(* CODESYS project listof.library
   DefaultNamespace: KOSTAL.AF2024.Core.ListOf
   DocFormat: reStructuredText
   Description: Lists of different elements
   Author: Frank Dümpelmann
   Title: KOSTAL.AF2024.Core.ListOf
   Version: 1.0.0.0
   Company: KOSTAL GmbH & Co.KG
   Placeholder: KOSTAL.AF2024.Core.ListOf

Project tree, tasks and I/O mapping:
  libraries: KOSTAL.AF2024.Core.functionResponse, 0.0.0.2 (KOSTAL GmbH & Co.KG); KOSTAL.AF2024.Core.Settings, 0.0.0.1 (KOSTAL GmbH & Co.KG); KOSTAL.AF2024.Core.System, 0.0.0.1 (KOSTAL GmbH & Co.KG); Tc2_Standard, 3.3.3.0 (Beckhoff Automation GmbH)
  _Interface/
    0_Core/
      BaseElement/
        data type _P_Interface
        data type _ST_Interface
      function block _FB_Interface_Core [ST]: FB_exit, FB_init, _addItem, _findItem, _findItemByIndex, _insertItem, _removeFromBegin, _removeFromEnd, _removeItem, _removeItemByIndex, _nextItem, _previousItem, _clearResult, _setResultFail, _setResultPass, _checkConsistency, _clear, _NumberOfMember, _RegKey
      interface _I_Interface_Core
      interface _I_Interface_Core_Owner
    1_Base/
      function block _FB_Interface_Base [ST]: _verifyMember, _addMember, _findMember, _findMemberByIndex, _insertMember, _removeFromBegin, _removeFromEnd, _removeMember, _removeMemberByIndex, _clear, FB_exit, FB_init
      interface _I_Interface_Base
      interface _I_Interface_Base_Owner
  _Object/
    function block _FB_Object_Base [ST]: _removePayload, _removeMember, _clear, FB_exit, FB_init
    interface _I_Object_Base
    interface _I_Object_Base_Owner
  _STRING/
    0_Core/
      BaseElement/
        data type _P_String
        data type _ST_String
      function block _FB_String_Core [ST]: _addItem, _findItem, _findItemByIndex, _insertItem, _removeFromBegin, _removeFromEnd, _removeItem, _removeItemByIndex, _nextItem, _previousItem, _clearResult, _setResultFail, _setResultPass, _checkConsistency, _clear, _NumberOfMember, FB_exit, FB_init
      interface _I_String_Core
      interface _I_String_Core_Owner
    1_Base/
      function block _FB_String_Base [ST]: _FIFO_peek, _FIFO_pop, _FIFO_push, _addMember, _findMember, _findMemberByIndex, _insertMember, _removeFromBegin, _removeFromEnd, _removeMember, _removeMemberByIndex, _clear, FB_exit, FB_init
      interface _I_String_Base
      interface _I_String_Base_Owner
    function block FB_ListOfString [ST]: addLine, clear, line_GET, line_SET, maxLine, NumberOfLines, removeLine
    interface I_ListOfString: line_GET, maxLine, NumberOfLines
    interface I_ListOfString_Owner: addLine, clear, line_GET, line_SET, maxLine, NumberOfLines, removeLine
  _STRING_UTF8/
    0_Core/
      BaseElement/
        data type P_String_UTF8
        data type ST_String_UTF8
      function block _FB_String_UTF8_Core [ST]: _addItem, _findItem, _findItemByIndex, _insertItem, _removeFromBegin, _removeFromEnd, _removeItem, _removeItemByIndex, _nextItem, _previousItem, _clearResult, _setResultFail, _setResultPass, _checkConsistency, _clear, _NumberOfMember, FB_exit, FB_init
      interface _I_String_UTF8_Core
      interface _I_String_UTF8_Core_Owner
    1_Base/
      function block _FB_String_UTF8_Base [ST]: _FIFO_peek, _FIFO_pop, _FIFO_push, _addMember, _findMember, _findMemberByIndex, _insertMember, _removeFromBegin, _removeFromEnd, _removeMember, _removeMemberByIndex, _clear, FB_exit, FB_init
      interface _I_String_UTF8_Base
      interface _I_String_UTF8_Base_Owner
    function block FB_ListOfString_UTF8 [ST]: addLine, clear, line_GET, line_SET, maxLine, NumberOfLines, removeLine
    interface I_ListOfString_UTF8: line_GET, maxLine, NumberOfLines
    interface I_ListOfString_UTF8_Owner: addLine, clear, line_GET, line_SET, maxLine, NumberOfLines, removeLine
  Project Information/
    function F_GetCompany [ST]
    function F_GetTitle [ST]
    function F_GetVersion [ST]
  Version/
    global variables Global_Version
*)

// _Interface/0_Core/BaseElement/_P_Interface
//Pointer to an element of List
TYPE _P_Interface : POINTER TO _ST_Interface; END_TYPE

// _Interface/0_Core/BaseElement/_ST_Interface
{attribute 'enable_dynamic_creation'}
TYPE _ST_Interface :
	STRUCT
			pNext	 		: _P_Interface;				//Pointer to next Item
			iMember		: KOSTAL_AF2024_Core_System.I_Interface;	//Interface of this item
			pPrevious : _P_Interface;				//Pointer to previous item
	END_STRUCT
END_TYPE

// _STRING/0_Core/BaseElement/_P_String
//Pointer to an element of List
TYPE _P_String : POINTER TO _ST_String; END_TYPE

// _STRING/0_Core/BaseElement/_ST_String
{attribute 'enable_dynamic_creation'}
TYPE _ST_String :
	STRUCT
			pNext	 		: _P_String;														//Pointer to next Item
			Member		: KOSTAL_AF2024_Core_Settings.T_MaxString;	//Text content
			pPrevious : _P_String;														//Pointer to previous item
	END_STRUCT
END_TYPE

// _STRING_UTF8/0_Core/BaseElement/P_String_UTF8
//Pointer to an element of List
TYPE P_String_UTF8 : POINTER TO ST_String_UTF8; END_TYPE

// _STRING_UTF8/0_Core/BaseElement/ST_String_UTF8
{attribute 'enable_dynamic_creation'}
TYPE ST_String_UTF8 :
	STRUCT
			pNext	 		: P_String_UTF8;				//Pointer to next Item
			Member			: KOSTAL_AF2024_Core_Settings.T_MaxString_UTF8;	//Text content
			pPrevious : P_String_UTF8;				//Pointer to previous item
	END_STRUCT
END_TYPE

// Version/Global_Version
{attribute 'TcGenerated'}
{attribute 'no-analysis'}
{attribute 'linkalways'}
// This function has been automatically generated from the project information.
VAR_GLOBAL CONSTANT
	{attribute 'const_non_replaced'}
	stLibVersion_KOSTAL_AF2024_Core_ListOf : ST_LibVersion := (iMajor := 1, iMinor := 0, iBuild := 0, iRevision := 0, nFlags := 0, sVersion := '1.0.0.0');
END_VAR

// _Interface/0_Core/_FB_Interface_Core
(*

| =========================================================================
| List of Items from base Interface {KOSTAL_TC3_Core_System.I_Interface} 
| =========================================================================

..code::

	//In addition to the interface, each item contains the pointer to the previous item 
	//as well as the pointer to the next item in the list.

	TYPE ST_List :
		STRUCT
				pNext			: P_List;
				iMember		: KOSTAL_TC3_Core_System.I_Interface;	
				pPrevious : P_List;
		END_STRUCT
	END_TYPE

============= ======================================= ======================
| The List is defined by (p)Begin and (p)End and also the count of Members 
----------------------------------------------------------------------------
============= ======================================= ======================
 **_pBegin**  >>>>>>>>>>>>>>>>>>>>>>>>>>>>>>>>>>>>>>  **_pEnd**                     
 **Item-1**	    Item-2   Item-3   Item-4  Item-5      **Item-n**                   
============= ======================================= ======================



| =========================================================================
| The Member is an Interface as payload and an access pointer to the        
| previous member and the next member                                      
| ---------------------------------------------------------------------------
| Previous Item ---<<<Pointer-Previous-[Item]-Pointer-Next>>>---NextItem---
| =========================================================================

*)
FUNCTION_BLOCK ABSTRACT _FB_Interface_Core IMPLEMENTS _I_Interface_Core, _I_Interface_Core_Owner

VAR
	_pBegin	: _P_Interface;	//origin of List
  _pEnd		: _P_Interface;	//end of List
	_Count	: UDINT;	//number of registered Member
	
	_RegKeyValue	: UDINT:= UDINT#0;	//use to create an unique ID
	
END_VAR

METHOD FB_exit : BOOL
VAR_INPUT
	bInCopyCode : BOOL; // if TRUE, the exit method is called for exiting an instance that is copied afterwards (online change).
END_VAR

_clear();
END_METHOD

METHOD FB_init : BOOL
VAR_INPUT
	bInitRetains : BOOL; // if TRUE, the retain variables are initialized (warm start / cold start)
	bInCopyCode : BOOL;  // if TRUE, the instance afterwards gets moved into the copy code (online change)
END_VAR

_clear();
END_METHOD

(*
	add new item to end of list
*)
METHOD PROTECTED _addItem : BOOL

VAR_INPUT
	Item		: KOSTAL_AF2024_Core_System.I_Interface;
	Result	: KOSTAL_AF2024_Core_functionResponse.I_T_functionResponse_Owner;
END_VAR

VAR
	_pNewItem	: _P_Interface;
END_VAR

_clearResult(Result);

IF Item = 0 THEN _setResultFail(Result, "Parameter Item is empty");	RETURN;	END_IF


//create a new Item
_pNewItem:= __NEW(_ST_Interface);

//If creation failed 
IF _pNewItem = 0 THEN _setResultFail(Result, "New Item cannot create");	RETURN;	END_IF

//If list is empty
IF THIS^._Count = 0 (*THIS^._pEnd = 0*) THEN THIS^._pBegin:= THIS^._pEnd:= _pNewItem; 
ELSE

	//set new item previous item to actual last item (THIS^._pEnd)
	_pNewItem^.pPrevious:= THIS^._pEnd;
	_pNewItem^.pPrevious^.pNext:= _pNewItem;
 
	THIS^._pEnd:= _pNewItem;
END_IF

THIS^._pEnd^.iMember:= Item;
THIS^._Count:= THIS^._Count + UDINT#1;

_setResultPass(Result, "addItem successful");

_RegKeyValue:= _RegKeyValue + 1;

_addItem:= TRUE;
END_METHOD

(*
	Search for the element {Item} in the list and return {FoundItem} if it is found {_findItem = TRUE}
*)
METHOD PROTECTED _findItem : BOOL
VAR_INPUT
	Item			: KOSTAL_AF2024_Core_System.I_Interface;
	FoundItem	: REFERENCE TO _P_Interface;
	Result		: KOSTAL_AF2024_Core_functionResponse.I_T_functionResponse_Owner;
END_VAR

VAR
	_Item		: _P_Interface;
END_VAR

_clearResult(Result);

IF Item = 0 										THEN _setResultFail(Result, "Parameter Item is empty");	RETURN;	END_IF
IF NOT __ISVALIDREF(FoundItem)	THEN _setResultFail(Result, "FoundItem has no valid reference");	RETURN;	END_IF


_Item := THIS^._pBegin;

WHILE _Item <> 0 DO

	IF _Item^.iMember = Item THEN

		FoundItem := _Item;

		_findItem:= TRUE;

		_setResultPass(Result, "Item found");
		
		RETURN;   

	END_IF
	
	_Item := THIS^._nextItem(_Item, 0);

END_WHILE

//FoundItem:= _Item;

_setResultFail(Result, "Item not found");

_findItem:= FALSE;
END_METHOD

(*
	Search for the element {Item} in the list and return {FoundItem} if it is found {_findItem = TRUE}
*)
METHOD PROTECTED _findItemByIndex : BOOL
VAR_INPUT
	Index			: UDINT;
	FoundItem	: REFERENCE TO _P_Interface;
	Result		: KOSTAL_AF2024_Core_functionResponse.I_T_functionResponse_Owner;
END_VAR

VAR
	_Item		: _P_Interface;
	_udi: UDINT;
END_VAR

_findItemByIndex:= FALSE;

_clearResult(Result);

IF _Count = 0										THEN _setResultFail(Result, "List is empty");											RETURN;	END_IF
IF Index > (_Count - 1)					THEN _setResultFail(Result, "Parameter Index is out of range");		RETURN;	END_IF
IF NOT __ISVALIDREF(FoundItem)	THEN _setResultFail(Result, "FoundItem has no valid reference");	RETURN;	END_IF

//set index 0
_Item := THIS^._pBegin;

//increase until index is reached
FOR _udi:= 1 TO Index DO
		_Item := THIS^._nextItem(_Item, 0);
END_FOR

FoundItem:= _Item;

IF FoundItem = 0 THEN
	_setResultFail(Result, "Item not found");
ELSE	
	_setResultPass(Result, "Item found");
	_findItemByIndex:= TRUE;
END_IF
END_METHOD

METHOD PROTECTED _insertItem : BOOL
VAR_INPUT
	Index		: UDINT;	//Index a which shall inserted the {Item}
	Item		: KOSTAL_AF2024_Core_System.I_Interface;
	Result		: KOSTAL_AF2024_Core_functionResponse.I_T_functionResponse_Owner;
END_VAR

VAR
	_pNewItem			: _P_Interface;
	_pExitingItem	: _P_Interface;
END_VAR

_clearResult(Result);

//Item is empty
IF Item = 0 THEN _setResultFail(Result, "Parameter Item is empty");	RETURN;	END_IF

//if List is empty add item 
IF (Index = 0) AND (_Count = 0)	THEN _insertItem:= _addItem(Item, Result);	RETURN;	END_IF

//Index is in list not available 
IF Index > (_Count - 1) THEN _setResultFail(Result, "Index is out of range");	RETURN;	END_IF

//if index is end of list then add item to end of list 
IF (Index = (_Count - 1)) THEN _insertItem:= _addItem(Item, Result);	RETURN;	END_IF

//try to find item where shall inserted
IF NOT _findItemByIndex(Index, _pExitingItem, Result) THEN RETURN;	END_IF
IF _pExitingItem = 0 THEN _setResultFail(Result, "Item not available");	RETURN;	END_IF


//create a new Item
_pNewItem:= __NEW(_ST_Interface);

//If creation failed 
IF _pNewItem = 0 THEN _setResultFail(Result, "New Item cannot create");	RETURN;	END_IF

_pNewItem^.iMember:= Item;

_pNewItem^.pNext		:= _pExitingItem;							//set the next item from new item to existing founded item
_pNewItem^.pPrevious:= _pExitingItem^.pPrevious;	//set the previous from existing item to the previous of new item

//if a previous exist then
//set the next from previous from existing item to the previous of new item
IF _pNewItem^.pPrevious <> 0 THEN	_pNewItem^.pPrevious^.pNext:= _pNewItem;	END_IF

_pExitingItem^.pPrevious:= _pNewItem;							//set the previous from existing founded item to  new item

//if inserted at the begin of list, set the begin pointer to new Item
IF _pBegin = _pExitingItem THEN	_pBegin:= _pNewItem;	END_IF

_Count:= _Count + UDINT#1;

_setResultPass(Result, "insertItem successful");

_RegKeyValue:= _RegKeyValue + 1;

_insertItem:= TRUE;
END_METHOD

(*
	remove Item from begin of list
*)
METHOD PROTECTED _removeFromBegin : BOOL
VAR_INPUT
	Result	: KOSTAL_AF2024_Core_functionResponse.I_T_functionResponse_Owner;
END_VAR

_removeFromBegin:= _removeItemByIndex(0, Result);
END_METHOD

(*
	remove Item from end of list
*)
METHOD PROTECTED _removeFromEnd : BOOL
VAR_INPUT
	Result	: KOSTAL_AF2024_Core_functionResponse.I_T_functionResponse_Owner;
END_VAR

_removeFromEnd:= _removeItemByIndex(_Count - 1, Result);
END_METHOD

(*
	remove given {Item} from List
*)
METHOD PROTECTED _removeItem : BOOL
VAR_INPUT
	Item		: _P_Interface;
	Result	: KOSTAL_AF2024_Core_functionResponse.I_T_functionResponse_Owner;
END_VAR

_clearResult(Result);

IF Item = 0 THEN _setResultFail(Result, "Parameter Item is empty");	RETURN;	END_IF

//exist a next member
IF Item^.pNext <> 0 THEN
	//set next members previous Item  to my previous Item
	Item^.pNext^.pPrevious := Item^.pPrevious; 
END_IF

//exist a previous member
IF Item^.pPrevious <> 0 THEN
	//set previous members next Item  to my next Item
	Item^.pPrevious^.pNext := Item^.pNext;
END_IF

//Item is the once member
IF Item = _pBegin AND Item = _pEnd THEN
	
	_pBegin := 0;
	_pEnd := 0;

ELSIF Item = _pBegin (*AND Item <> THIS^._pEnd*) THEN

	_pBegin := Item^.pNext;

ELSIF Item = _pEnd THEN

	_pEnd := Item^.pPrevious;

END_IF

__DELETE(Item);

IF  _Count > UDINT#0 THEN	_Count := _Count - UDINT#1;	
ELSE
	_setResultFail(Result, "removeItem Counter underflow");
	RETURN;
END_IF

_setResultPass(Result, "removeItem successful");
_removeItem:= TRUE;
END_METHOD

(*
	remove given {Index} from List
*)
METHOD PROTECTED _removeItemByIndex : BOOL
VAR_INPUT
	Index		: UDINT;
	Result	: KOSTAL_AF2024_Core_functionResponse.I_T_functionResponse_Owner;
END_VAR

VAR
	_Item		: _P_Interface;
	_bFound	: BOOL;
END_VAR

IF NOT _findItemByIndex(Index, _Item, Result)	THEN RETURN;	END_IF

_removeItemByIndex:= _removeItem(_Item, Result);
END_METHOD

// retreives the pointer to the next item of the given entry
METHOD PROTECTED _nextItem : _P_Interface;
VAR_INPUT
    Item : _P_Interface;
		Result	: KOSTAL_AF2024_Core_functionResponse.I_T_functionResponse_Owner;
END_VAR
VAR
	_Res	: _P_Interface;
END_VAR

IF Item <> 0 THEN	_Res := Item^.pNext;
ELSE							_Res := 0;
END_IF

_nextItem:= _Res;
END_METHOD

// retreives the previous item of the given entry
METHOD PROTECTED _previousItem : _P_Interface
VAR_INPUT
    Item 	: _P_Interface;
END_VAR
VAR
	_Res	: _P_Interface;
END_VAR

IF Item <> 0 THEN	_Res := Item^.pPrevious;
ELSE							_Res := 0;
END_IF

_previousItem:= _Res;
END_METHOD

(*
	Clear result component
*)
METHOD PROTECTED _clearResult : BOOL
VAR_INPUT
	IN : KOSTAL_AF2024_Core_functionResponse.I_T_functionResponse_Owner;
END_VAR

IF IN <> 0 THEN  
	 IN.clear();
	_clearResult:= TRUE;	
END_IF
END_METHOD

(*
	set result to fail with given information 
*)
METHOD PROTECTED _setResultFail : BOOL
VAR_INPUT
	IN 		: KOSTAL_AF2024_Core_functionResponse.I_T_functionResponse_Owner;
	Info	: KOSTAL_AF2024_Core_Settings.T_MaxString;
END_VAR

IF IN <> 0 THEN 

	IN.success:= FALSE;
	IN.status:= Info;

	_setResultFail:= TRUE;

END_IF
END_METHOD

(*
	set result to pass with given information 
*)
METHOD PROTECTED _setResultPass : BOOL
VAR_INPUT
	IN 		: KOSTAL_AF2024_Core_functionResponse.I_T_functionResponse_Owner;
	Info	: KOSTAL_AF2024_Core_Settings.T_MaxString;
END_VAR

IF IN <> 0 THEN 

	IN.success:= TRUE;
	IN.status:= Info;

	_setResultPass:= TRUE;

END_IF
END_METHOD

(*
	Check if the list is consistent
*)
METHOD PROTECTED _checkConsistency : BOOL
VAR_INPUT
	Result	: KOSTAL_AF2024_Core_functionResponse.I_T_functionResponse_Owner;
END_VAR

VAR
	_pItem			: _P_Interface;
	_pNext			: _P_Interface;
	_pPrev			: _P_Interface;
	_nItemCounter	: UDINT;
	_bBeginOk			: BOOL;
	_bEndOk			: BOOL;
	_bPrevLinkOk		: BOOL;
	_bNextLinkOk		: BOOL;
	_bItemCountOk	: BOOL;
	_bInterfaceOk	: BOOL;
END_VAR

// check from pHead to pTail
_pItem:= _pBegin;
_nItemCounter:= 0;

IF _pBegin <> 0 THEN
	_bBeginOk:= (_pBegin^.pPrevious = 0);
ELSE
	_bBeginOk:= TRUE;
END_IF

IF _pEnd <> 0 THEN
	_bEndOk:= (_pEnd^.pNext = 0);
ELSE
	_bEndOk:= TRUE;
END_IF

IF _bBeginOk AND _bEndOk THEN

	_bPrevLinkOk:= TRUE;
	_bNextLinkOk:= TRUE;
	_bInterfaceOk:= TRUE;

	WHILE _pItem <> 0 DO
		
		_pPrev:= _pItem^.pPrevious;
		_pNext:= _pItem^.pNext;

		IF _pPrev <> 0 THEN
			_bPrevLinkOk:= (_pPrev^.pNext = _pItem);
		ELSE
			_bPrevLinkOk:= (_pItem = _pBegin);
		END_IF

		IF _pNext <> 0 THEN
			_bNextLinkOk:= (_pNext^.pPrevious = _pItem);
		ELSE
			_bNextLinkOk:= (_pItem = _pEnd);
		END_IF

		_bInterfaceOk:= (_pItem^.iMember <> 0);

		IF NOT _bNextLinkOk OR NOT _bPrevLinkOk OR NOT _bInterfaceOk THEN	EXIT;	END_IF

		//handle iteration
		_nItemCounter:= _nItemCounter + UDINT#1;
		_pItem:= _nextItem(_pItem, 0);

	END_WHILE

END_IF

_bItemCountOk:= (_nItemCounter = THIS^._Count);

IF 		NOT _bBeginOk			THEN	_setResultFail(Result, "List head not ok");
ELSIF NOT _bEndOk				THEN	_setResultFail(Result, "List End not ok");
ELSIF NOT _bPrevLinkOk 	THEN	_setResultFail(Result, Tc2_Standard.WCONCAT("Previous Link failed by item ", UDINT_TO_WSTRING(_nItemCounter)));
ELSIF NOT _bNextLinkOk	THEN	_setResultFail(Result, Tc2_Standard.WCONCAT("Next Link failed by item ", UDINT_TO_WSTRING(_nItemCounter)));
ELSIF NOT	_bInterfaceOk	THEN	_setResultFail(Result, Tc2_Standard.WCONCAT("Interface failed by item ", UDINT_TO_WSTRING(_nItemCounter))); 
ELSIF NOT	_bItemCountOk THEN	_setResultFail(Result, "Itemcounter is not ok");
ELSE													_setResultPass(Result, "List is consistent");	_checkConsistency:= TRUE;
END_IF
END_METHOD

(*
	Delete the complete content of the list
*)
METHOD PROTECTED _clear

WHILE THIS^._pBegin <> 0 DO
    THIS^._removeItem(THIS^._pBegin, 0);  
END_WHILE
END_METHOD

//return the nnumber of items in List
PROPERTY PROTECTED _NumberOfMember : UDINT
GET

_NumberOfMember:= _Count;
END_GET
END_PROPERTY

PROPERTY PROTECTED _RegKey : UDINT
GET

_RegKey:= THIS^._RegKeyValue;
END_GET
END_PROPERTY

END_FUNCTION_BLOCK

// _Interface/0_Core/_I_Interface_Core
INTERFACE _I_Interface_Core EXTENDS KOSTAL_AF2024_Core_System.I_Interface

END_INTERFACE

// _Interface/0_Core/_I_Interface_Core_Owner
INTERFACE _I_Interface_Core_Owner EXTENDS KOSTAL_AF2024_Core_System.I_Interface

END_INTERFACE

// _Interface/1_Base/_FB_Interface_Base
(*

| =========================================================================
| List of Items from base Interface {KOSTAL_TC3_Core_System.I_Interface} 
| =========================================================================

..code::

	//In addition to the interface, each item contains the pointer to the previous item 
	//as well as the pointer to the next item in the list.

	TYPE ST_List :
		STRUCT
				pNext			: P_List;
				iMember		: KOSTAL_TC3_Core_System.I_Interface;	
				pPrevious : P_List;
		END_STRUCT
	END_TYPE

============= ======================================= ======================
| The List is defined by (p)Begin and (p)End and also the count of Members 
----------------------------------------------------------------------------
============= ======================================= ======================
 **_pBegin**  >>>>>>>>>>>>>>>>>>>>>>>>>>>>>>>>>>>>>>  **_pEnd**                     
 **Item-1**	    Item-2   Item-3   Item-4  Item-5      **Item-n**                   
============= ======================================= ======================



| =========================================================================
| The Member is an Interface as payload and an access pointer to the        
| previous member and the next member                                      
| ---------------------------------------------------------------------------
| Previous Item ---<<<Pointer-Previous-[Item]-Pointer-Next>>>---NextItem---
| =========================================================================

*)
FUNCTION_BLOCK ABSTRACT _FB_Interface_Base EXTENDS _FB_Interface_Core IMPLEMENTS _I_Interface_Base, _I_Interface_Base_Owner

(*
	integrate here the veryfing of your interface type 
	only if verifing is passed [_verifyMember:= TRUE] the called metode will proceeded 
*)
METHOD PROTECTED _verifyMember : BOOL

VAR_INPUT
	Member	: KOSTAL_AF2024_Core_System.I_Interface;
	Result	: KOSTAL_AF2024_Core_functionResponse.I_T_functionResponse_Owner;
END_VAR

VAR
	_obj	: KOSTAL_AF2024_Core_System.I_Interface;
	_bResult: BOOL;
END_VAR

IF Member = 0 THEN _setResultFail(Result, "Parameter Member is empty");	RETURN;	END_IF

_bResult:= __QUERYINTERFACE(Member, _obj);

IF NOT _bResult OR (_obj = 0) THEN
	IF Result <> 0 THEN  
		Result.success:= FALSE; 
		Result.status:= "no valid interface found";	
	END_IF	
	RETURN;
END_IF

_verifyMember:= TRUE;
END_METHOD

(*
	add new Member to end of list
*)
METHOD PROTECTED _addMember : BOOL

VAR_INPUT
	Member		: KOSTAL_AF2024_Core_System.I_Interface;
	Result	: KOSTAL_AF2024_Core_functionResponse.I_T_functionResponse_Owner;
END_VAR


VAR
	_Member: KOSTAL_AF2024_Core_System.I_Interface;
END_VAR

//IF NOT _verifyMember(Member, Result)	THEN	RETURN;	END_IF

//member already exist
IF _findMember(Member,_Member, Result) THEN 
	_setResultFail(Result, "The participant already exists in the list.");
	RETURN;	
END_IF	

_addMember:= _addItem(Member, Result);
END_METHOD

(*
	Search for the element {Item} in the list and return {FoundItem} if it is found {_findItem = TRUE}
*)
METHOD PROTECTED _findMember : BOOL
VAR_INPUT
	Member			: KOSTAL_AF2024_Core_System.I_Interface;
	FoundMember	: REFERENCE TO KOSTAL_AF2024_Core_System.I_Interface;	//return value
	Result			: KOSTAL_AF2024_Core_functionResponse.I_T_functionResponse_Owner;
END_VAR

VAR
	_Item		: _P_Interface;
END_VAR

_clearResult(Result);

IF Member = 0 												THEN _setResultFail(Result, "Parameter Item is empty");	RETURN;	END_IF
IF NOT __ISVALIDREF(FoundMember)			THEN _setResultFail(Result, "FoundItem has no valid reference");	RETURN;	END_IF
IF NOT _verifyMember(Member, Result)	THEN	RETURN;	END_IF

_findMember:= _findItem(Member, _Item, Result);

IF NOT _findMember		THEN	RETURN;	END_IF
IF _Item = 0 					THEN	RETURN;	END_IF
//IF _Item^.iMember = 0 THEN	RETURN;	END_IF
IF NOT _verifyMember(_Item^.iMember, Result)	THEN	RETURN;	END_IF

FoundMember:= _Item^.iMember;
END_METHOD

//find a modul by index  
METHOD PROTECTED _findMemberByIndex : BOOL
VAR_INPUT
	Index				: UDINT;	//index of item
	FoundMember	: REFERENCE TO KOSTAL_AF2024_Core_System.I_Interface;	//return value
	Result			: KOSTAL_AF2024_Core_functionResponse.I_T_functionResponse_Owner;	//result information
END_VAR

VAR
	_FoundItem	: _P_Interface;
END_VAR

IF NOT __ISVALIDREF(FoundMember)	THEN _setResultFail(Result, "FoundMember has no valid reference");	RETURN;	END_IF

FoundMember:= 0;

_findMemberByIndex:= _findItemByIndex(Index,_FoundItem, Result);

IF NOT _findMemberByIndex THEN RETURN;	END_IF

IF NOT _verifyMember(_FoundItem^.iMember, Result) THEN RETURN;	END_IF

FoundMember:= _FoundItem^.iMember;

_findMemberByIndex:= TRUE;
END_METHOD

METHOD PROTECTED _insertMember : BOOL
VAR_INPUT
	Index		: UDINT;	//Index a which shall inserted the {Item}
	Member	: KOSTAL_AF2024_Core_System.I_Interface;
	Result	:KOSTAL_AF2024_Core_functionResponse.I_T_functionResponse_Owner;
END_VAR

VAR
	_Member: KOSTAL_AF2024_Core_System.I_Interface;
END_VAR

//IF NOT _verifyMember(Member, Result)	THEN	RETURN;	END_IF

//member already exist
IF _findMember(Member,_Member, Result) THEN 
	_setResultFail(Result, "The participant already exists in the list.");
	RETURN;	
END_IF	

_insertMember:= _insertItem(Index, Member, Result);
END_METHOD

(*
	remove Item from begin of list
*)
METHOD PROTECTED _removeFromBegin : BOOL
VAR_INPUT
	Result	: KOSTAL_AF2024_Core_functionResponse.I_T_functionResponse_Owner;
END_VAR

_removeFromBegin:= _removeMemberByIndex(0, Result);
END_METHOD

(*
	remove Item from end of list
*)
METHOD PROTECTED _removeFromEnd : BOOL
VAR_INPUT
	Result	: KOSTAL_AF2024_Core_functionResponse.I_T_functionResponse_Owner;
END_VAR

_removeFromEnd:= _removeMemberByIndex(_Count - 1, Result);
END_METHOD

(*
	remove given {Member} from List
*)
METHOD PROTECTED _removeMember : BOOL
VAR_INPUT
	Member	: KOSTAL_AF2024_Core_System.I_Interface;
	Result	: KOSTAL_AF2024_Core_functionResponse.I_T_functionResponse_Owner;
END_VAR

VAR
	_Item		: _P_Interface;
	_bFound: BOOL;
END_VAR


IF NOT _verifyMember(Member, Result)	THEN	RETURN;	END_IF

_bFound:= _findItem(Member, _Item, Result);

IF NOT _bFound THEN RETURN;	END_IF

_removeMember:= _removeItem(_Item, Result);
END_METHOD

(*
	remove given {Index} from List
*)
METHOD PROTECTED _removeMemberByIndex : BOOL
VAR_INPUT
	Index		: UDINT;
	Result	: KOSTAL_AF2024_Core_functionResponse.I_T_functionResponse_Owner;
END_VAR

VAR
	_bFound	: BOOL;
	_Member	: KOSTAL_AF2024_Core_System.I_Interface;

END_VAR

IF NOT _findMemberByIndex(Index, _Member, Result)	THEN RETURN;	END_IF

_removeMemberByIndex:= _removeMember(_Member, Result);
END_METHOD

(*
	Delete the complete content of the list
*)
METHOD PROTECTED _clear
VAR_INPUT
END_VAR

WHILE THIS^._pBegin <> 0 DO
    THIS^._removeMember(THIS^._pBegin^.iMember, 0);  
END_WHILE
END_METHOD

METHOD FB_exit : BOOL
VAR_INPUT
	bInCopyCode : BOOL; // if TRUE, the exit method is called for exiting an instance that is copied afterwards (online change).
END_VAR

_clear();
END_METHOD

METHOD FB_init : BOOL
VAR_INPUT
	bInitRetains : BOOL; // if TRUE, the retain variables are initialized (warm start / cold start)
	bInCopyCode : BOOL;  // if TRUE, the instance afterwards gets moved into the copy code (online change)
END_VAR

_clear();
END_METHOD

END_FUNCTION_BLOCK

// _Interface/1_Base/_I_Interface_Base
INTERFACE _I_Interface_Base EXTENDS _I_Interface_Core

END_INTERFACE

// _Interface/1_Base/_I_Interface_Base_Owner
INTERFACE _I_Interface_Base_Owner EXTENDS _I_Interface_Core_Owner

END_INTERFACE

// _Object/_FB_Object_Base
(*

| ==================================================================================
| List of Items of objects with base Interface {KOSTAL_TC3_Core_System.I_Interface} 
| ==================================================================================

..code::

	//In addition to the interface, each item contains the pointer to the previous item 
	//as well as the pointer to the next item in the list.

	TYPE ST_List :
		STRUCT
				pNext			: P_List;
				iMember		: KOSTAL_TC3_Core_System.I_Interface;	
				pPrevious : P_List;
		END_STRUCT
	END_TYPE

============= ======================================= ======================
| The List is defined by (p)Begin and (p)End and also the count of Members 
----------------------------------------------------------------------------
============= ======================================= ======================
 **_pBegin**  >>>>>>>>>>>>>>>>>>>>>>>>>>>>>>>>>>>>>>  **_pEnd**                     
 **Item-1**	    Item-2   Item-3   Item-4  Item-5      **Item-n**                   
============= ======================================= ======================



| =========================================================================
| The Member is an object which implements the base Interface as payload. 
| -------------------------------------------------------------------------
| Previous Item ---<<<Pointer-Previous-[Item]-Pointer-Next>>>---NextItem---
| =========================================================================

*)
FUNCTION_BLOCK ABSTRACT _FB_Object_Base EXTENDS _FB_Interface_Base IMPLEMENTS _I_Object_Base, _I_Object_Base_Owner

(*
	Integrate the type-specific procedures here to clean up the member and remove it from memory. 
	only if verifing is passed [_verifyMember:= TRUE] the called metode should proceed 
*)
METHOD PROTECTED _removePayload : BOOL
VAR_INPUT
	Member	: KOSTAL_AF2024_Core_System.I_Interface;
	Result	: KOSTAL_AF2024_Core_functionResponse.I_T_functionResponse_Owner;
END_VAR

_removePayload:= TRUE;
END_METHOD

(*
	remove given {Member} from List including the customer payload {_removePayload()]
*)
METHOD PROTECTED _removeMember : BOOL
VAR_INPUT
	Member	: KOSTAL_AF2024_Core_System.I_Interface;
	Result	: KOSTAL_AF2024_Core_functionResponse.I_T_functionResponse_Owner;
END_VAR

VAR
	_Item		: _P_Interface;
	_bFound: BOOL;
END_VAR

IF NOT _verifyMember(Member, Result)	THEN	RETURN;	END_IF

_bFound:= _findItem(Member, _Item, Result);

IF NOT _bFound THEN RETURN;	END_IF

_removePayload(Member, Result);

_removeMember:= _removeItem(_Item, Result);
END_METHOD

(*
	Delete the complete content of the list including the customer payload {_removePayload()}
*)
METHOD PROTECTED _clear

WHILE THIS^._pBegin <> 0 DO
  _removeMember(_pBegin^.iMember, 0);  
END_WHILE
END_METHOD

METHOD FB_exit : BOOL
VAR_INPUT
	bInCopyCode : BOOL; // if TRUE, the exit method is called for exiting an instance that is copied afterwards (online change).
END_VAR

_clear();
END_METHOD

METHOD FB_init : BOOL
VAR_INPUT
	bInitRetains : BOOL; // if TRUE, the retain variables are initialized (warm start / cold start)
	bInCopyCode : BOOL;  // if TRUE, the instance afterwards gets moved into the copy code (online change)
END_VAR

_clear();
END_METHOD

END_FUNCTION_BLOCK

// _Object/_I_Object_Base
INTERFACE _I_Object_Base EXTENDS _I_Interface_Base

END_INTERFACE

// _Object/_I_Object_Base_Owner
INTERFACE _I_Object_Base_Owner EXTENDS _I_Interface_Base_Owner

END_INTERFACE

// _STRING/0_Core/_FB_String_Core
(*

| =========================================================================
| List of Items from base Interface {KOSTAL_TC3_Core_System.I_Interface} 
| =========================================================================

..code::

	//In addition to the interface, each item contains the pointer to the previous item 
	//as well as the pointer to the next item in the list.

	TYPE ST_List :
		STRUCT
				pNext			: P_List;
				iMember		: KOSTAL_TC3_Core_System.I_Interface;	
				pPrevious : P_List;
		END_STRUCT
	END_TYPE

============= ======================================= ======================
| The List is defined by (p)Begin and (p)End and also the count of Members 
----------------------------------------------------------------------------
============= ======================================= ======================
 **_pBegin**  >>>>>>>>>>>>>>>>>>>>>>>>>>>>>>>>>>>>>>  **_pEnd**                     
 **Item-1**	    Item-2   Item-3   Item-4  Item-5      **Item-n**                   
============= ======================================= ======================



| =========================================================================
| The Member is an Interface as payload and an access pointer to the        
| previous member and the next member                                      
| ---------------------------------------------------------------------------
| Previous Item ---<<<Pointer-Previous-[Item]-Pointer-Next>>>---NextItem---
| =========================================================================

*)
FUNCTION_BLOCK ABSTRACT _FB_String_Core IMPLEMENTS _I_String_Core, _I_String_Core_Owner

VAR
	_pBegin	: _P_String;	//origin of List
  _pEnd		: _P_String;	//end of List
	_Count	: UDINT;	//number of registered Member
END_VAR

(*
	add new item to end of list
*)
METHOD PROTECTED _addItem : BOOL

VAR_INPUT
	Member	: KOSTAL_AF2024_Core_Settings.T_MaxString;
	Result	: KOSTAL_AF2024_Core_functionResponse.I_T_functionResponse_Owner;
END_VAR

VAR
	_pNewItem	: _P_String;
END_VAR

_clearResult(Result);

//IF Item = 0 THEN _setResultFail(Result, 'Parameter Item is empty');	RETURN;	END_IF


//create a new Item
_pNewItem:= __NEW(_ST_String);

//If creation failed 
IF _pNewItem = 0 THEN _setResultFail(Result, "New Item cannot create");	RETURN;	END_IF

//If list is empty
IF _Count = 0 THEN _pBegin:= _pEnd:= _pNewItem; 
ELSE

	//set new item previous item to actual last item (THIS^._pEnd)
	_pNewItem^.pPrevious:= _pEnd;
	_pNewItem^.pPrevious^.pNext:= _pNewItem;
 
	_pEnd:= _pNewItem;

END_IF

_pEnd^.Member:= Member;
_Count:= _Count + UDINT#1;

_setResultPass(Result, "addItem successful");

_addItem:= TRUE;
END_METHOD

(*
	Search for the element {Item} in the list and return {FoundItem} if it is found {_findItem = TRUE}
*)
METHOD PROTECTED _findItem : BOOL
VAR_INPUT
	Member		: KOSTAL_AF2024_Core_Settings.T_MaxString;
	FoundItem	: REFERENCE TO _P_String;
	Result		: KOSTAL_AF2024_Core_functionResponse.I_T_functionResponse_Owner;
END_VAR

VAR
	_Item		: _P_String;
END_VAR

_clearResult(Result);

IF NOT __ISVALIDREF(FoundItem)	THEN _setResultFail(Result, "FoundItem has no valid reference");	RETURN;	END_IF


_Item := _pBegin;

WHILE _Item <> 0 DO

	IF _Item^.Member = Member THEN

		FoundItem := _Item;

		_findItem:= TRUE;

		_setResultPass(Result, "Item found");
		
		RETURN;   

	END_IF
	
	_Item := _nextItem(_Item, 0);

END_WHILE

//FoundItem:= _Item;

_setResultFail(Result, "Item not found");

_findItem:= FALSE;
END_METHOD

(*
	Search for the element {Item} in the list and return {FoundItem} if it is found {_findItem = TRUE}
*)
METHOD PROTECTED _findItemByIndex : BOOL
VAR_INPUT
	Index			: UDINT;
	FoundItem	: REFERENCE TO _P_String;
	Result		: KOSTAL_AF2024_Core_functionResponse.I_T_functionResponse_Owner;
END_VAR

VAR
	_Item	: _P_String;
	_udi	: UDINT;
END_VAR

_findItemByIndex:= FALSE;

_clearResult(Result);

IF _Count = 0										THEN _setResultFail(Result, "List is empty");											RETURN;	END_IF
IF Index > (_Count - 1)					THEN _setResultFail(Result, "Parameter Index is out of range");		RETURN;	END_IF
IF NOT __ISVALIDREF(FoundItem)	THEN _setResultFail(Result, "FoundItem has no valid reference");	RETURN;	END_IF


_Item := _pBegin;

FOR _udi:= 1 TO Index DO
		_Item := _nextItem(_Item, 0);
END_FOR

FoundItem:= _Item;

IF FoundItem = 0 THEN
	_setResultFail(Result, "Item not found");
ELSE	
	_setResultPass(Result, "Item found");
	_findItemByIndex:= TRUE;
END_IF
END_METHOD

METHOD PROTECTED _insertItem : BOOL
VAR_INPUT
	Index		: UDINT;	//Index a which shall inserted the {Item}
	Member	: KOSTAL_AF2024_Core_Settings.T_MaxString;
	Result	: KOSTAL_AF2024_Core_functionResponse.I_T_functionResponse_Owner;
END_VAR

VAR
	_pNewItem			: _P_String;
	_pExitingItem	: _P_String;
END_VAR
_clearResult(Result);

//if List is empty add item 
IF (Index = 0) AND (_Count = 0)	THEN _insertItem:= _addItem(Member, Result);	RETURN;	END_IF

//Index is in list not available 
IF Index > (_Count - 1) THEN _setResultFail(Result, "Index is out of range");	RETURN;	END_IF

//if index is end of list then add item to end of list 
IF (Index = (_Count - 1)) THEN _insertItem:= _addItem(Member, Result);	RETURN;	END_IF

//try to find item where shall inserted
IF NOT _findItemByIndex(Index, _pExitingItem, Result) THEN RETURN;	END_IF
IF _pExitingItem = 0 THEN _setResultFail(Result, "Item not available");	RETURN;	END_IF


//create a new Item
_pNewItem:= __NEW(_ST_String);

//If creation failed 
IF _pNewItem = 0 THEN _setResultFail(Result, "New Item cannot create");	RETURN;	END_IF

_pNewItem^.Member:= Member;

_pNewItem^.pNext		:= _pExitingItem;							//set the next item from new item to existing founded item
_pNewItem^.pPrevious:= _pExitingItem^.pPrevious;	//set the previous from existing item to the previous of new item

//if a previous exist then
//set the next from previous from existing item to the previous of new item
IF _pNewItem^.pPrevious <> 0 THEN	_pNewItem^.pPrevious^.pNext:= _pNewItem;	END_IF

_pExitingItem^.pPrevious:= _pNewItem;							//set the previous from existing founded item to  new item

//if inserted at the begin of list, set the begin pointer to new Item
IF _pBegin = _pExitingItem THEN	_pBegin:= _pNewItem;	END_IF

_Count:= _Count + UDINT#1;

_setResultPass(Result, "insertItem successful");

_insertItem:= TRUE;
END_METHOD

(*
	remove Item from begin of list
*)
METHOD PROTECTED _removeFromBegin : BOOL
VAR_INPUT
	Result	: KOSTAL_AF2024_Core_functionResponse.I_T_functionResponse_Owner;
END_VAR

_removeFromBegin:= _removeItemByIndex(0, Result);
END_METHOD

(*
	remove Item from end of list
*)
METHOD PROTECTED _removeFromEnd : BOOL
VAR_INPUT
	Result	: KOSTAL_AF2024_Core_functionResponse.I_T_functionResponse_Owner;
END_VAR

_removeFromEnd:= _removeItemByIndex(_Count - 1, Result);
END_METHOD

(*
	remove given {Item} from List
*)
METHOD PROTECTED _removeItem : BOOL
VAR_INPUT
	Item		: _P_String;
	Result	: KOSTAL_AF2024_Core_functionResponse.I_T_functionResponse_Owner;
END_VAR

_clearResult(Result);

IF Item = 0 THEN _setResultFail(Result, "Parameter Item is empty");	RETURN;	END_IF

//exist a next member
IF Item^.pNext <> 0 THEN
	//set next members previous Item  to my previous Item
	Item^.pNext^.pPrevious := Item^.pPrevious; 
END_IF

//exist a previous member
IF Item^.pPrevious <> 0 THEN
	//set previous members next Item  to my next Item
	Item^.pPrevious^.pNext := Item^.pNext;
END_IF

//Item is the once member
IF Item = _pBegin AND Item = _pEnd THEN
	
	_pBegin := 0;
	_pEnd := 0;

ELSIF Item = _pBegin THEN

	_pBegin := Item^.pNext;

ELSIF Item = _pEnd THEN

	_pEnd := Item^.pPrevious;

END_IF

__DELETE(Item);

IF  _Count > UDINT#0 THEN	_Count := _Count - UDINT#1;	
ELSE
	_setResultFail(Result, "removeItem Counter underflow");
	RETURN;
END_IF

_setResultPass(Result, "removeItem successful");
_removeItem:= TRUE;
END_METHOD

(*
	remove given {Index} from List
*)
METHOD PROTECTED _removeItemByIndex : BOOL
VAR_INPUT
	Index		: UDINT;
	Result	: KOSTAL_AF2024_Core_functionResponse.I_T_functionResponse_Owner;
END_VAR

VAR
	_Item		: _P_String;
	_bFound	: BOOL;
END_VAR

IF NOT _findItemByIndex(Index, _Item, Result)	THEN RETURN;	END_IF

_removeItemByIndex:= _removeItem(_Item, Result);
END_METHOD

// retreives the pointer to the next item of the given entry
METHOD PROTECTED _nextItem : _P_String;
VAR_INPUT
    Item : _P_String;
		Result	: KOSTAL_AF2024_Core_functionResponse.I_T_functionResponse_Owner;
END_VAR
VAR
	_Res	: _P_String;
END_VAR

IF Item <> 0 THEN	_Res := Item^.pNext;
ELSE							_Res := 0;
END_IF

_nextItem:= _Res;
END_METHOD

// retreives the previous item of the given entry
METHOD PROTECTED _previousItem : _P_String
VAR_INPUT
    Item 	: _P_String;
END_VAR
VAR
	_Res	: _P_String;
END_VAR

IF Item <> 0 THEN	_Res := Item^.pPrevious;
ELSE							_Res := 0;
END_IF

_previousItem:= _Res;
END_METHOD

(*
	Clear result component
*)
METHOD PROTECTED _clearResult : BOOL
VAR_INPUT
	IN : KOSTAL_AF2024_Core_functionResponse.I_T_functionResponse_Owner;
END_VAR

IF IN <> 0 THEN 
	IN.clear(); 
	_clearResult:= TRUE;	
END_IF
END_METHOD

(*
	set result to fail with given information 
*)
METHOD PROTECTED _setResultFail : BOOL
VAR_INPUT
	IN 		: KOSTAL_AF2024_Core_functionResponse.I_T_functionResponse_Owner;
	Info	: KOSTAL_AF2024_Core_Settings.T_MaxString;
END_VAR

IF IN <> 0 THEN 

	IN.success:= FALSE;
	IN.status:= Info;

	_setResultFail:= TRUE;

END_IF
END_METHOD

(*
	set result to pass with given information 
*)
METHOD PROTECTED _setResultPass : BOOL
VAR_INPUT
	IN 		: KOSTAL_AF2024_Core_functionResponse.I_T_functionResponse_Owner;
	Info	: KOSTAL_AF2024_Core_Settings.T_MaxString;
END_VAR

IF IN <> 0 THEN 

	IN.success:= TRUE;
	IN.status:= Info;

	_setResultPass:= TRUE;

END_IF
END_METHOD

(*
	Check if the list is consistent
*)
METHOD PROTECTED _checkConsistency : BOOL
VAR_INPUT
	Result	: KOSTAL_AF2024_Core_functionResponse.I_T_functionResponse_Owner;
END_VAR

VAR
	_pItem			: _P_String;
	_pNext			: _P_String;
	_pPrev			: _P_String;
	_nItemCounter	: UDINT;
	_bBeginOk			: BOOL;
	_bEndOk			: BOOL;
	_bPrevLinkOk		: BOOL;
	_bNextLinkOk		: BOOL;
	_bItemCountOk	: BOOL;
END_VAR
// check from pHead to pTail
_pItem:= _pBegin;
_nItemCounter:= 0;

IF _pBegin <> 0 THEN
	_bBeginOk:= (_pBegin^.pPrevious = 0);
ELSE
	_bBeginOk:= TRUE;
END_IF

IF _pEnd <> 0 THEN
	_bEndOk:= (_pEnd^.pNext = 0);
ELSE
	_bEndOk:= TRUE;
END_IF

IF _bBeginOk AND _bEndOk THEN

	_bPrevLinkOk:= TRUE;
	_bNextLinkOk:= TRUE;

	WHILE _pItem <> 0 DO
		
		_pPrev:= _pItem^.pPrevious;
		_pNext:= _pItem^.pNext;

		IF _pPrev <> 0 THEN
			_bPrevLinkOk:= (_pPrev^.pNext = _pItem);
		ELSE
			_bPrevLinkOk:= (_pItem = _pBegin);
		END_IF

		IF _pNext <> 0 THEN
			_bNextLinkOk:= (_pNext^.pPrevious = _pItem);
		ELSE
			_bNextLinkOk:= (_pItem = THIS^._pEnd);
		END_IF

		IF NOT _bNextLinkOk OR NOT _bPrevLinkOk THEN	EXIT;	END_IF

		//handle iteration
		_nItemCounter:= _nItemCounter + UDINT#1;
		_pItem:= _nextItem(_pItem, 0);

	END_WHILE

END_IF

_bItemCountOk:= (_nItemCounter = THIS^._Count);

IF 		NOT _bBeginOk			THEN	_setResultFail(Result, "List head not ok");
ELSIF NOT _bEndOk				THEN	_setResultFail(Result, "List End not ok");
ELSIF NOT _bPrevLinkOk 	THEN	_setResultFail(Result, Tc2_Standard.WCONCAT("Previous Link failed by item ", UDINT_TO_WSTRING(_nItemCounter)));
ELSIF NOT _bNextLinkOk	THEN	_setResultFail(Result, Tc2_Standard.WCONCAT("Next Link failed by item ", UDINT_TO_WSTRING(_nItemCounter)));
ELSIF NOT	_bItemCountOk THEN	_setResultFail(Result, "Itemcounter is not ok");
ELSE													_setResultPass(Result, "List is consistent");	_checkConsistency:= TRUE;
END_IF
END_METHOD

(*
	Delete the complete content of the list
*)
METHOD PROTECTED _clear

WHILE THIS^._pBegin <> 0 DO
  _removeItem(_pBegin, 0);  
END_WHILE
END_METHOD

//return the nnumber of items in List
PROPERTY PROTECTED _NumberOfMember : UDINT
GET

_NumberOfMember:= _Count;
END_GET
END_PROPERTY

METHOD FB_exit : BOOL
VAR_INPUT
	bInCopyCode : BOOL; // if TRUE, the exit method is called for exiting an instance that is copied afterwards (online change).
END_VAR

_clear();
END_METHOD

METHOD FB_init : BOOL
VAR_INPUT
	bInitRetains : BOOL; // if TRUE, the retain variables are initialized (warm start / cold start)
	bInCopyCode : BOOL;  // if TRUE, the instance afterwards gets moved into the copy code (online change)
END_VAR

_clear();
END_METHOD

END_FUNCTION_BLOCK

// _STRING/0_Core/_I_String_Core
INTERFACE _I_String_Core EXTENDS KOSTAL_AF2024_Core_System.I_Interface

END_INTERFACE

// _STRING/0_Core/_I_String_Core_Owner
INTERFACE _I_String_Core_Owner EXTENDS KOSTAL_AF2024_Core_System.I_Interface

END_INTERFACE

// _STRING/1_Base/_FB_String_Base
(*

| =========================================================================
| List of Items from base Interface {KOSTAL_TC3_Core_System.I_Interface} 
| =========================================================================

..code::

	//In addition to the interface, each item contains the pointer to the previous item 
	//as well as the pointer to the next item in the list.

	TYPE ST_List :
		STRUCT
				pNext			: P_List;
				Line			: KOSTAL_TC3_Core_Settings.T_MaxString;	//Text content
				pPrevious : P_List;
		END_STRUCT
	END_TYPE

============= ======================================= ======================
| The List is defined by (p)Begin and (p)End and also the count of Members 
----------------------------------------------------------------------------
============= ======================================= ======================
 **_pBegin**  >>>>>>>>>>>>>>>>>>>>>>>>>>>>>>>>>>>>>>  **_pEnd**                     
 **Item-1**	    Item-2   Item-3   Item-4  Item-5      **Item-n**                   
============= ======================================= ======================



| =========================================================================
| The Member is an Interface as payload and an access pointer to the        
| previous member and the next member                                      
| ---------------------------------------------------------------------------
| Previous Item ---<<<Pointer-Previous-[Item]-Pointer-Next>>>---NextItem---
| =========================================================================

*)
FUNCTION_BLOCK ABSTRACT _FB_String_Base EXTENDS _FB_String_Core IMPLEMENTS _I_String_Base, _I_String_Base_Owner

//methode return the Member from begin 
METHOD PROTECTED _FIFO_peek : BOOL
VAR_INPUT
	FoundMember	: REFERENCE TO KOSTAL_AF2024_Core_Settings.T_MaxString;	//return value
	Result			: KOSTAL_AF2024_Core_functionResponse.I_T_functionResponse_Owner;
END_VAR

_clearResult(Result);

IF 		NOT __ISVALIDREF(FoundMember) THEN _setResultFail(Result, "FoundMember has no valid reference"); 
ELSE	_FIFO_peek:= _findMemberByIndex(0, FoundMember, Result);
END_IF
END_METHOD

//methode return the Member from begin and remove it from List
METHOD PROTECTED _FIFO_pop : BOOL
VAR_INPUT
	FoundMember	: REFERENCE TO KOSTAL_AF2024_Core_Settings.T_MaxString;	//return value
	Result			: KOSTAL_AF2024_Core_functionResponse.I_T_functionResponse_Owner;
END_VAR


_clearResult(Result);

_FIFO_pop:= _findMemberByIndex(0, FoundMember, Result);

IF _FIFO_pop THEN	_FIFO_pop:= _removeFromBegin(Result);	END_IF
END_METHOD

//push/add the {Member} to begin from List
METHOD PROTECTED _FIFO_push : BOOL
VAR_INPUT
	Member	: KOSTAL_AF2024_Core_Settings.T_MaxString;
	Result	: KOSTAL_AF2024_Core_functionResponse.I_T_functionResponse_Owner;
END_VAR


_FIFO_push:= _addItem(Member, Result);
END_METHOD

(*
	add new Member to end of list
*)
METHOD PROTECTED _addMember : BOOL

VAR_INPUT
	Member		: KOSTAL_AF2024_Core_Settings.T_MaxString;
	Result	: KOSTAL_AF2024_Core_functionResponse.I_T_functionResponse_Owner;
END_VAR


VAR
	_Member: KOSTAL_AF2024_Core_System.I_Interface;
END_VAR

_addMember:= _addItem(Member, Result);
END_METHOD

(*
	Search for the element {Item} in the list and return {FoundItem} if it is found {_findItem = TRUE}
*)
METHOD PROTECTED _findMember : BOOL
VAR_INPUT
	Member			: KOSTAL_AF2024_Core_Settings.T_MaxString;
	FoundMember	: REFERENCE TO KOSTAL_AF2024_Core_Settings.T_MaxString;	//return value
	Result			: KOSTAL_AF2024_Core_functionResponse.I_T_functionResponse_Owner;
END_VAR

VAR
	_Item		: _P_String;
END_VAR

_clearResult(Result);

IF NOT __ISVALIDREF(FoundMember) THEN _setResultFail(Result, "FoundItem has no valid reference");	RETURN;	END_IF

_findMember:= _findItem(Member, _Item, Result);

IF NOT _findMember		THEN	RETURN;	END_IF
IF _Item = 0 					THEN	RETURN;	END_IF

FoundMember:= _Item^.Member;
END_METHOD

//find a modul by index  
METHOD PROTECTED _findMemberByIndex : BOOL
VAR_INPUT
	Index				: UDINT;	//index of item
	FoundMember	: REFERENCE TO KOSTAL_AF2024_Core_Settings.T_MaxString;	//return value
	Result			: KOSTAL_AF2024_Core_functionResponse.I_T_functionResponse_Owner;	//result information
END_VAR

VAR
	_FoundItem	: _P_String;
END_VAR

IF NOT __ISVALIDREF(FoundMember)	THEN _setResultFail(Result, "FoundMember has no valid reference");	RETURN;	END_IF

FoundMember:= "";

_findMemberByIndex:= _findItemByIndex(Index,_FoundItem, Result);

IF NOT _findMemberByIndex	THEN RETURN;	END_IF
IF _FoundItem = 0 				THEN RETURN;	END_IF

FoundMember:= _FoundItem^.Member;

_findMemberByIndex:= TRUE;
END_METHOD

METHOD PROTECTED _insertMember : BOOL
VAR_INPUT
	Index		: UDINT;	//Index a which shall inserted the {Item}
	Member	: KOSTAL_AF2024_Core_Settings.T_MaxString;
	Result	: KOSTAL_AF2024_Core_functionResponse.I_T_functionResponse_Owner;
END_VAR

_insertMember:= _insertItem(Index, Member, Result);
END_METHOD

(*
	remove Item from begin of list
*)
METHOD PROTECTED _removeFromBegin : BOOL
VAR_INPUT
	Result	: KOSTAL_AF2024_Core_functionResponse.I_T_functionResponse_Owner;
END_VAR

_removeFromBegin:= _removeMemberByIndex(0, Result);
END_METHOD

(*
	remove Item from end of list
*)
METHOD PROTECTED _removeFromEnd : BOOL
VAR_INPUT
	Result	: KOSTAL_AF2024_Core_functionResponse.I_T_functionResponse_Owner;
END_VAR

_removeFromEnd:= _removeMemberByIndex(_Count - 1, Result);
END_METHOD

(*
	remove given {Member} from List
*)
METHOD PROTECTED _removeMember : BOOL
VAR_INPUT
	Member	: KOSTAL_AF2024_Core_Settings.T_MaxString;
	Result	: KOSTAL_AF2024_Core_functionResponse.I_T_functionResponse_Owner;
END_VAR

VAR
	_Item		: _P_String;
	_bFound: BOOL;
END_VAR


_bFound:= _findItem(Member, _Item, Result);

IF NOT _bFound THEN RETURN;	END_IF

_removeMember:= _removeItem(_Item, Result);
END_METHOD

(*
	remove given {Index} from List
*)
METHOD PROTECTED _removeMemberByIndex : BOOL
VAR_INPUT
	Index		: UDINT;
	Result	: KOSTAL_AF2024_Core_functionResponse.I_T_functionResponse_Owner;
END_VAR

VAR
	_bFound	: BOOL;
	_Member	: KOSTAL_AF2024_Core_Settings.T_MaxString;

END_VAR

IF NOT _findMemberByIndex(Index, _Member, Result)	THEN RETURN;	END_IF

_removeMemberByIndex:= _removeMember(_Member, Result);
END_METHOD

(*
	Delete the complete content of the list
*)
METHOD PROTECTED _clear
VAR_INPUT
END_VAR

WHILE THIS^._pBegin <> 0 DO
    _removeMember(_pBegin^.Member, 0);  
END_WHILE
END_METHOD

METHOD FB_exit : BOOL
VAR_INPUT
	bInCopyCode : BOOL; // if TRUE, the exit method is called for exiting an instance that is copied afterwards (online change).
END_VAR

_clear();
END_METHOD

METHOD FB_init : BOOL
VAR_INPUT
	bInitRetains : BOOL; // if TRUE, the retain variables are initialized (warm start / cold start)
	bInCopyCode : BOOL;  // if TRUE, the instance afterwards gets moved into the copy code (online change)
END_VAR

_clear();
END_METHOD

END_FUNCTION_BLOCK

// _STRING/1_Base/_I_String_Base
INTERFACE _I_String_Base EXTENDS _I_String_Core

END_INTERFACE

// _STRING/1_Base/_I_String_Base_Owner
INTERFACE _I_String_Base_Owner EXTENDS _I_String_Core_Owner

END_INTERFACE

// _STRING/FB_ListOfString
(*
	List of String
	HP -High Performance
	The temporary load on the router's memory is halved.
*)
FUNCTION_BLOCK PUBLIC FB_ListOfString EXTENDS _FB_String_Base IMPLEMENTS I_ListOfString, I_ListOfString_Owner
VAR
	_maxLine	: UDINT:= UDINT#16#FFFF_FFFF;
END_VAR

(*
Description
===========
| Adds a line to end of the list
| Parameters:
| 	line: STRING(255): Text to add to the list
| Returns false in case line is empty or list is full
*)
METHOD addLine : BOOL
VAR_INPUT
	newLine	: KOSTAL_AF2024_Core_Settings.T_MaxString;
END_VAR

VAR
	_fRes: KOSTAL_AF2024_Core_functionResponse.T_functionResponse;
END_VAR

addLine:= _addMember(newLine, _fRes) AND _fRes.success;
END_METHOD

(*
Description
===========
| Clears the list's contents
*)
METHOD clear

_clear();
END_METHOD

(*
Description
===========
| Returns the line at the given index
| Parameters:
| 	numberOfLine: index
*)
METHOD line_GET : KOSTAL_AF2024_Core_Settings.T_MaxString
VAR_INPUT
	(*1..numberOfLines_GET()*)
	numberOfLine	: UDINT;
END_VAR

VAR
	_fRes: KOSTAL_AF2024_Core_functionResponse.T_functionResponse;
END_VAR

_findMemberByIndex(NumberOfLine - 1, line_GET, _fRes);
END_METHOD

(*
Description
===========
| Returns the line at the given index
| Parameters:
| 	numberOfLine: index
*)
METHOD line_SET : BOOL
VAR_INPUT
	line	: KOSTAL_AF2024_Core_Settings.T_MaxString;
	(*1..numberOfLines_GET()*)
	numberOfLine	: UDINT;
END_VAR

VAR
	_item: _P_String;
	_fRes: KOSTAL_AF2024_Core_functionResponse.T_functionResponse;
END_VAR

IF NOT _findItemByIndex(numberOfLine - 1, _item, _fRes)	THEN RETURN;	END_IF

IF NOT _fRes.success	THEN RETURN;	END_IF

IF _item = 0 THEN RETURN;	END_IF

_item^.Member:= line;

line_SET:= TRUE;
END_METHOD

(*
Description
===========
| **Maximum** number of elements in the list. 
| If the list is full, added lines will be ignored
*)
PROPERTY maxLine : UDINT
GET

maxLine:= _maxLine;
END_GET
SET

_maxLine:= maxLine;
END_SET
END_PROPERTY

PROPERTY PUBLIC NumberOfLines : UDINT
GET

NumberOfLines:= SUPER^._Count;
END_GET
END_PROPERTY

(*
Description
===========
| Remove the line with the given index
| Elements after the index move up one position
| Parameters:
| 	index: line to remove
*)
METHOD removeLine
VAR_INPUT
	(*1..numberOfLines_GET()*)
	numberOfLine	: UDINT;
END_VAR

VAR
	_fRes: KOSTAL_AF2024_Core_functionResponse.T_functionResponse;
END_VAR

_removeMemberByIndex(numberOfLine - 1, _fRes);
END_METHOD

END_FUNCTION_BLOCK

// _STRING/I_ListOfString
INTERFACE I_ListOfString EXTENDS _I_String_Base

(*
Description
===========
| Returns the line at the given index
| Parameters:
| 	numberOfLine: index
*)
METHOD PUBLIC line_GET : KOSTAL_AF2024_Core_Settings.T_MaxString
VAR_INPUT
	numberOfLine	:	UDINT;	//1..numberOfLines_GET()
END_VAR
END_METHOD

(*
Description
===========
| **Maximum** number of elements in the list. 
| If the list is full, added lines will be ignored
*)
PROPERTY PUBLIC maxLine : UDINT
GET
END_GET
END_PROPERTY

PROPERTY PUBLIC NumberOfLines : UDINT
GET
END_GET
END_PROPERTY

END_INTERFACE

// _STRING/I_ListOfString_Owner
INTERFACE I_ListOfString_Owner EXTENDS _I_String_Base_Owner

(*
Description
===========
| Adds a line to end of the list
| Parameters:
| 	line: STRING(255): Text to add to the list
| Returns false in case line is empty or list is full
*)

METHOD PUBLIC addLine : BOOL
VAR_INPUT
	newLine	: KOSTAL_AF2024_Core_Settings.T_MaxString;
END_VAR
END_METHOD

(*
Description
===========
| Clears the list's contents
*)
METHOD PUBLIC clear
VAR_INPUT
END_VAR
END_METHOD

(*
Description
===========
| Returns the line at the given index
| Parameters:
| 	numberOfLine: index
*)
METHOD PUBLIC line_GET : KOSTAL_AF2024_Core_Settings.T_MaxString
VAR_INPUT
	numberOfLine	:	UDINT;	//1..numberOfLines_GET()
END_VAR
END_METHOD

(*
Description
===========
| Returns the line at the given index
| Parameters:
| 	numberOfLine: index
*)
METHOD PUBLIC line_SET : BOOL
VAR_INPUT
	line					: KOSTAL_AF2024_Core_Settings.T_MaxString;
	numberOfLine	:	UDINT;	//1..numberOfLines_GET()
END_VAR
END_METHOD

(*
Description
===========
| **Maximum** number of elements in the list. 
| If the list is full, added lines will be ignored
*)
PROPERTY PUBLIC maxLine : UDINT
GET
END_GET
SET
END_SET
END_PROPERTY

PROPERTY PUBLIC NumberOfLines : UDINT
GET
END_GET
END_PROPERTY

(*
Description
===========
| Remove the line with the given index
| Elements after the index move up one position
| Parameters:
| 	index: line to remove
*)

METHOD PUBLIC removeLine
VAR_INPUT
	numberOfLine	:	UDINT;	//1..numberOfLines_GET()
END_VAR
END_METHOD

END_INTERFACE

// _STRING_UTF8/0_Core/_FB_String_UTF8_Core
(*

| =========================================================================
| List of Items from base Interface {KOSTAL_AF2024_Core_System.I_Interface} 
| =========================================================================

..code::

	//In addition to the interface, each item contains the pointer to the previous item 
	//as well as the pointer to the next item in the list.

	TYPE ST_List :
		STRUCT
				pNext			: P_List;
				iMember		: KOSTAL_AF2024_Core_System.I_Interface;	
				pPrevious : P_List;
		END_STRUCT
	END_TYPE

============= ======================================= ======================
| The List is defined by (p)Begin and (p)End and also the count of Members 
----------------------------------------------------------------------------
============= ======================================= ======================
 **_pBegin**  >>>>>>>>>>>>>>>>>>>>>>>>>>>>>>>>>>>>>>  **_pEnd**                     
 **Item-1**	    Item-2   Item-3   Item-4  Item-5      **Item-n**                   
============= ======================================= ======================



| =========================================================================
| The Member is an Interface as payload and an access pointer to the        
| previous member and the next member                                      
| ---------------------------------------------------------------------------
| Previous Item ---<<<Pointer-Previous-[Item]-Pointer-Next>>>---NextItem---
| =========================================================================

*)
FUNCTION_BLOCK ABSTRACT _FB_String_UTF8_Core IMPLEMENTS _I_String_UTF8_Core, _I_String_UTF8_Core_Owner

VAR
	_pBegin	: P_String_UTF8;	//origin of List
  _pEnd		: P_String_UTF8;	//end of List
	_Count	: UDINT;	//number of registered Member
END_VAR

(*
	add new item to end of list
*)
METHOD PROTECTED _addItem : BOOL

VAR_INPUT
	Member		: KOSTAL_AF2024_Core_Settings.T_MaxString_UTF8;
	Result	: KOSTAL_AF2024_Core_functionResponse.I_T_functionResponse_Owner;
END_VAR

VAR
	_pNewItem	: P_String_UTF8;
END_VAR

_clearResult(Result);

//IF Item = 0 THEN _setResultFail(Result, 'Parameter Item is empty');	RETURN;	END_IF


//create a new Item
_pNewItem:= __NEW(ST_String_UTF8);

//If creation failed 
IF _pNewItem = 0 THEN _setResultFail(Result, "New Item cannot create");	RETURN;	END_IF

//If list is empty
IF _Count = 0 THEN _pBegin:= _pEnd:= _pNewItem; 
ELSE

	//set new item previous item to actual last item (THIS^._pEnd)
	_pNewItem^.pPrevious:= _pEnd;
	_pNewItem^.pPrevious^.pNext:= _pNewItem;
 
	_pEnd:= _pNewItem;
END_IF

_pEnd^.Member:= Member;
_Count:= _Count + UDINT#1;

_setResultPass(Result, "addItem successful");

_addItem:= TRUE;
END_METHOD

(*
	Search for the element {Item} in the list and return {FoundItem} if it is found {_findItem = TRUE}
*)
METHOD PROTECTED _findItem : BOOL
VAR_INPUT
	Member		: KOSTAL_AF2024_Core_Settings.T_MaxString_UTF8;
	FoundItem	: REFERENCE TO P_String_UTF8;
	Result		: KOSTAL_AF2024_Core_functionResponse.I_T_functionResponse_Owner;
END_VAR

VAR
	_Item		: P_String_UTF8;
END_VAR

_clearResult(Result);

IF NOT __ISVALIDREF(FoundItem)	THEN _setResultFail(Result, "FoundItem has no valid reference");	RETURN;	END_IF


_Item := _pBegin;

WHILE _Item <> 0 DO

	IF _Item^.Member = Member THEN

		FoundItem := _Item;

		_findItem:= TRUE;

		_setResultPass(Result, "Item found");
		
		RETURN;   

	END_IF
	
	_Item := _nextItem(_Item, 0);

END_WHILE

//FoundItem:= _Item;

_setResultFail(Result, "Item not found");

_findItem:= FALSE;
END_METHOD

(*
	Search for the element {Item} in the list and return {FoundItem} if it is found {_findItem = TRUE}
*)
METHOD PROTECTED _findItemByIndex : BOOL
VAR_INPUT
	Index			: UDINT;
	FoundItem	: REFERENCE TO P_String_UTF8;
	Result		: KOSTAL_AF2024_Core_functionResponse.I_T_functionResponse_Owner;
END_VAR

VAR
	_Item		: P_String_UTF8;
	_udi: UDINT;
END_VAR

_findItemByIndex:= FALSE;

_clearResult(Result);

IF _Count = 0										THEN _setResultFail(Result, "List is empty");											RETURN;	END_IF
IF Index > (_Count - 1)					THEN _setResultFail(Result, "Parameter Index is out of range");		RETURN;	END_IF
IF NOT __ISVALIDREF(FoundItem)	THEN _setResultFail(Result, "FoundItem has no valid reference");	RETURN;	END_IF


_Item := _pBegin;

FOR _udi:= 1 TO Index DO
		_Item := _nextItem(_Item, 0);
END_FOR

FoundItem:= _Item;

IF FoundItem = 0 THEN
	_setResultFail(Result, "Item not found");
ELSE	
	_setResultPass(Result, "Item found");
	_findItemByIndex:= TRUE;
END_IF
END_METHOD

METHOD PROTECTED _insertItem : BOOL
VAR_INPUT
	Index		: UDINT;	//Index a which shall inserted the {Item}
	Member	: KOSTAL_AF2024_Core_Settings.T_MaxString_UTF8;
	Result	: KOSTAL_AF2024_Core_functionResponse.I_T_functionResponse_Owner;
END_VAR

VAR
	_pNewItem			: P_String_UTF8;
	_pExitingItem	: P_String_UTF8;
END_VAR
_clearResult(Result);

//if List is empty add item 
IF (Index = 0) AND (_Count = 0)	THEN _insertItem:= _addItem(Member, Result);	RETURN;	END_IF

//Index is in list not available 
IF Index > (_Count - 1) THEN _setResultFail(Result, "Index is out of range");	RETURN;	END_IF

//if index is end of list then add item to end of list 
IF (Index = (_Count - 1)) THEN _insertItem:= _addItem(Member, Result);	RETURN;	END_IF

//try to find item where shall inserted
IF NOT _findItemByIndex(Index, _pExitingItem, Result) THEN RETURN;	END_IF
IF _pExitingItem = 0 THEN _setResultFail(Result, "Item not available");	RETURN;	END_IF


//create a new Item
_pNewItem:= __NEW(ST_String_UTF8);

//If creation failed 
IF _pNewItem = 0 THEN _setResultFail(Result, "New Item cannot create");	RETURN;	END_IF

_pNewItem^.Member:= Member;

_pNewItem^.pNext		:= _pExitingItem;							//set the next item from new item to existing founded item
_pNewItem^.pPrevious:= _pExitingItem^.pPrevious;	//set the previous from existing item to the previous of new item

//if a previous exist then
//set the next from previous from existing item to the previous of new item
IF _pNewItem^.pPrevious <> 0 THEN	_pNewItem^.pPrevious^.pNext:= _pNewItem;	END_IF

_pExitingItem^.pPrevious:= _pNewItem;							//set the previous from existing founded item to  new item

//if inserted at the begin of list, set the begin pointer to new Item
IF _pBegin = _pExitingItem THEN	_pBegin:= _pNewItem;	END_IF

_Count:= _Count + UDINT#1;

_setResultPass(Result, "insertItem successful");

_insertItem:= TRUE;
END_METHOD

(*
	remove Item from begin of list
*)
METHOD PROTECTED _removeFromBegin : BOOL
VAR_INPUT
	Result	: KOSTAL_AF2024_Core_functionResponse.I_T_functionResponse_Owner;
END_VAR

_removeFromBegin:= _removeItemByIndex(0, Result);
END_METHOD

(*
	remove Item from end of list
*)
METHOD PROTECTED _removeFromEnd : BOOL
VAR_INPUT
	Result	: KOSTAL_AF2024_Core_functionResponse.I_T_functionResponse_Owner;
END_VAR

_removeFromEnd:= _removeItemByIndex(_Count - 1, Result);
END_METHOD

(*
	remove given {Item} from List
*)
METHOD PROTECTED _removeItem : BOOL
VAR_INPUT
	Item		: P_String_UTF8;
	Result	: KOSTAL_AF2024_Core_functionResponse.I_T_functionResponse_Owner;
END_VAR

_clearResult(Result);

IF Item = 0 THEN _setResultFail(Result, "Parameter Item is empty");	RETURN;	END_IF

//exist a next member
IF Item^.pNext <> 0 THEN
	//set next members previous Item  to my previous Item
	Item^.pNext^.pPrevious := Item^.pPrevious; 
END_IF

//exist a previous member
IF Item^.pPrevious <> 0 THEN
	//set previous members next Item  to my next Item
	Item^.pPrevious^.pNext := Item^.pNext;
END_IF

//Item is the once member
IF Item = _pBegin AND Item = _pEnd THEN
	
	_pBegin := 0;
	_pEnd := 0;

ELSIF Item = _pBegin THEN

	_pBegin := Item^.pNext;

ELSIF Item = _pEnd THEN

	_pEnd := Item^.pPrevious;

END_IF

__DELETE(Item);

IF  _Count > UDINT#0 THEN	_Count := _Count - UDINT#1;	
ELSE
	_setResultFail(Result, "removeItem Counter underflow");
	RETURN;
END_IF

_setResultPass(Result, "removeItem successful");
_removeItem:= TRUE;
END_METHOD

(*
	remove given {Index} from List
*)
METHOD PROTECTED _removeItemByIndex : BOOL
VAR_INPUT
	Index		: UDINT;
	Result	: KOSTAL_AF2024_Core_functionResponse.I_T_functionResponse_Owner;
END_VAR

VAR
	_Item		: P_String_UTF8;
	_bFound	: BOOL;
END_VAR

IF NOT _findItemByIndex(Index, _Item, Result)	THEN RETURN;	END_IF

_removeItemByIndex:= _removeItem(_Item, Result);
END_METHOD

// retreives the pointer to the next item of the given entry
METHOD PROTECTED _nextItem : P_String_UTF8;
VAR_INPUT
    Item : P_String_UTF8;
		Result	: KOSTAL_AF2024_Core_functionResponse.I_T_functionResponse_Owner;
END_VAR
VAR
	_Res	: P_String_UTF8;
END_VAR

IF Item <> 0 THEN	_Res := Item^.pNext;
ELSE							_Res := 0;
END_IF

_nextItem:= _Res;
END_METHOD

// retreives the previous item of the given entry
METHOD PROTECTED _previousItem : P_String_UTF8
VAR_INPUT
    Item 	: P_String_UTF8;
END_VAR
VAR
	_Res	: P_String_UTF8;
END_VAR

IF Item <> 0 THEN	_Res := Item^.pPrevious;
ELSE							_Res := 0;
END_IF

_previousItem:= _Res;
END_METHOD

(*
	Clear result component
*)
METHOD PROTECTED _clearResult : BOOL
VAR_INPUT
	IN : KOSTAL_AF2024_Core_functionResponse.I_T_functionResponse_Owner;
END_VAR

IF IN <> 0 THEN 
	IN.clear(); 
	_clearResult:= TRUE;	
END_IF
END_METHOD

(*
	set result to fail with given information 
*)
METHOD PROTECTED _setResultFail : BOOL
VAR_INPUT
	IN 		: KOSTAL_AF2024_Core_functionResponse.I_T_functionResponse_Owner;
	Info	: KOSTAL_AF2024_Core_Settings.T_MaxString;
END_VAR

IF IN <> 0 THEN 

	IN.success:= FALSE;
	IN.status:= Info;

	_setResultFail:= TRUE;

END_IF
END_METHOD

(*
	set result to pass with given information 
*)
METHOD PROTECTED _setResultPass : BOOL
VAR_INPUT
	IN 		: KOSTAL_AF2024_Core_functionResponse.I_T_functionResponse_Owner;
	Info	: KOSTAL_AF2024_Core_Settings.T_MaxString;
END_VAR

IF IN <> 0 THEN 

	IN.success:= TRUE;
	IN.status:= Info;

	_setResultPass:= TRUE;

END_IF
END_METHOD

(*
	Check if the list is consistent
*)
METHOD PROTECTED _checkConsistency : BOOL
VAR_INPUT
	Result	: KOSTAL_AF2024_Core_functionResponse.I_T_functionResponse_Owner;
END_VAR

VAR
	_pItem			: P_String_UTF8;
	_pNext			: P_String_UTF8;
	_pPrev			: P_String_UTF8;
	_nItemCounter	: UDINT;
	_bBeginOk			: BOOL;
	_bEndOk			: BOOL;
	_bPrevLinkOk		: BOOL;
	_bNextLinkOk		: BOOL;
	_bItemCountOk	: BOOL;
END_VAR
// check from pHead to pTail
_pItem:= _pBegin;
_nItemCounter:= 0;

IF _pBegin <> 0 THEN
	_bBeginOk:= (_pBegin^.pPrevious = 0);
ELSE
	_bBeginOk:= TRUE;
END_IF

IF _pEnd <> 0 THEN
	_bEndOk:= (_pEnd^.pNext = 0);
ELSE
	_bEndOk:= TRUE;
END_IF

IF _bBeginOk AND _bEndOk THEN

	_bPrevLinkOk:= TRUE;
	_bNextLinkOk:= TRUE;

	WHILE _pItem <> 0 DO
		
		_pPrev:= _pItem^.pPrevious;
		_pNext:= _pItem^.pNext;

		IF _pPrev <> 0 THEN
			_bPrevLinkOk:= (_pPrev^.pNext = _pItem);
		ELSE
			_bPrevLinkOk:= (_pItem = _pBegin);
		END_IF

		IF _pNext <> 0 THEN
			_bNextLinkOk:= (_pNext^.pPrevious = _pItem);
		ELSE
			_bNextLinkOk:= (_pItem = _pEnd);
		END_IF

		IF NOT _bNextLinkOk OR NOT _bPrevLinkOk THEN	EXIT;	END_IF

		//handle iteration
		_nItemCounter:= _nItemCounter + UDINT#1;
		_pItem:= _nextItem(_pItem, 0);

	END_WHILE

END_IF

_bItemCountOk:= (_nItemCounter = _Count);

IF 		NOT _bBeginOk			THEN	_setResultFail(Result, "List head not ok");
ELSIF NOT _bEndOk				THEN	_setResultFail(Result, "List End not ok");
ELSIF NOT _bPrevLinkOk 	THEN	_setResultFail(Result, Tc2_Standard.WCONCAT("Previous Link failed by item ", UDINT_TO_WSTRING(_nItemCounter)));
ELSIF NOT _bNextLinkOk	THEN	_setResultFail(Result, Tc2_Standard.WCONCAT("Next Link failed by item ", UDINT_TO_WSTRING(_nItemCounter)));
ELSIF NOT	_bItemCountOk THEN	_setResultFail(Result, "Itemcounter is not ok");
ELSE													_setResultPass(Result, "List is consistent");	_checkConsistency:= TRUE;
END_IF
END_METHOD

(*
	Delete the complete content of the list
*)
METHOD PROTECTED _clear

WHILE THIS^._pBegin <> 0 DO
	_removeItem(_pBegin, 0);  
END_WHILE
END_METHOD

//return the nnumber of items in List
PROPERTY PROTECTED _NumberOfMember : UDINT
GET

_NumberOfMember:= _Count;
END_GET
END_PROPERTY

METHOD FB_exit : BOOL
VAR_INPUT
	bInCopyCode : BOOL; // if TRUE, the exit method is called for exiting an instance that is copied afterwards (online change).
END_VAR

_clear();
END_METHOD

METHOD FB_init : BOOL
VAR_INPUT
	bInitRetains : BOOL; // if TRUE, the retain variables are initialized (warm start / cold start)
	bInCopyCode : BOOL;  // if TRUE, the instance afterwards gets moved into the copy code (online change)
END_VAR

_clear();
END_METHOD

END_FUNCTION_BLOCK

// _STRING_UTF8/0_Core/_I_String_UTF8_Core
INTERFACE _I_String_UTF8_Core EXTENDS KOSTAL_AF2024_Core_System.I_Interface

END_INTERFACE

// _STRING_UTF8/0_Core/_I_String_UTF8_Core_Owner
INTERFACE _I_String_UTF8_Core_Owner EXTENDS KOSTAL_AF2024_Core_System.I_Interface

END_INTERFACE

// _STRING_UTF8/1_Base/_FB_String_UTF8_Base
(*

| =========================================================================
| List of Items from base Interface {KOSTAL_AF2024_Core_System.I_Interface} 
| =========================================================================

..code::

	//In addition to the interface, each item contains the pointer to the previous item 
	//as well as the pointer to the next item in the list.

	TYPE ST_List :
		STRUCT
				pNext			: P_List;
				Line			: KOSTAL_AF2024_Core_Settings.T_MaxString_UTF8;	//Text content
				pPrevious : P_List;
		END_STRUCT
	END_TYPE

============= ======================================= ======================
| The List is defined by (p)Begin and (p)End and also the count of Members 
----------------------------------------------------------------------------
============= ======================================= ======================
 **_pBegin**  >>>>>>>>>>>>>>>>>>>>>>>>>>>>>>>>>>>>>>  **_pEnd**                     
 **Item-1**	    Item-2   Item-3   Item-4  Item-5      **Item-n**                   
============= ======================================= ======================



| =========================================================================
| The Member is an Interface as payload and an access pointer to the        
| previous member and the next member                                      
| ---------------------------------------------------------------------------
| Previous Item ---<<<Pointer-Previous-[Item]-Pointer-Next>>>---NextItem---
| =========================================================================

*)
FUNCTION_BLOCK ABSTRACT _FB_String_UTF8_Base EXTENDS _FB_String_UTF8_Core IMPLEMENTS _I_String_UTF8_Base, _I_String_UTF8_Base_Owner

VAR
END_VAR

//methode return the Member from begin 
METHOD PROTECTED _FIFO_peek : BOOL
VAR_INPUT
	FoundMember	: REFERENCE TO KOSTAL_AF2024_Core_Settings.T_MaxString_UTF8;	//return value
	Result			: KOSTAL_AF2024_Core_functionResponse.I_T_functionResponse_Owner;
END_VAR

_clearResult(Result);

IF 		NOT __ISVALIDREF(FoundMember) THEN _setResultFail(Result, "FoundMember has no valid reference"); 
ELSE	_FIFO_peek:= _findMemberByIndex(0, FoundMember, Result);
END_IF
END_METHOD

//methode return the Member from begin and remove it from List
METHOD PROTECTED _FIFO_pop : BOOL
VAR_INPUT
	FoundMember	: REFERENCE TO KOSTAL_AF2024_Core_Settings.T_MaxString_UTF8;	//return value
	Result			: KOSTAL_AF2024_Core_functionResponse.I_T_functionResponse_Owner;
END_VAR


_clearResult(Result);

_FIFO_pop:= _findMemberByIndex(0, FoundMember, Result);

IF _FIFO_pop THEN	_FIFO_pop:= _removeFromBegin(Result);	END_IF
END_METHOD

//push/add the {Member} to begin from List
METHOD PROTECTED _FIFO_push : BOOL
VAR_INPUT
	Member	: KOSTAL_AF2024_Core_Settings.T_MaxString_UTF8;
	Result	: KOSTAL_AF2024_Core_functionResponse.I_T_functionResponse_Owner;
END_VAR


_FIFO_push:= _addItem(Member, Result);
END_METHOD

(*
	add new Member to end of list
*)
METHOD PROTECTED _addMember : BOOL

VAR_INPUT
	Member		: KOSTAL_AF2024_Core_Settings.T_MaxString_UTF8;
	Result	: KOSTAL_AF2024_Core_functionResponse.I_T_functionResponse_Owner;
END_VAR


VAR
	_Member: KOSTAL_AF2024_Core_System.I_Interface;
END_VAR

_addMember:= _addItem(Member, Result);
END_METHOD

(*
	Search for the element {Item} in the list and return {FoundItem} if it is found {_findItem = TRUE}
*)
METHOD PROTECTED _findMember : BOOL
VAR_INPUT
	Member			: KOSTAL_AF2024_Core_Settings.T_MaxString_UTF8;
	FoundMember	: REFERENCE TO KOSTAL_AF2024_Core_Settings.T_MaxString_UTF8;	//return value
	Result			: KOSTAL_AF2024_Core_functionResponse.I_T_functionResponse_Owner;
END_VAR

VAR
	_Item		: P_String_UTF8;
END_VAR

_clearResult(Result);

IF NOT __ISVALIDREF(FoundMember)			THEN _setResultFail(Result, "FoundItem has no valid reference");	RETURN;	END_IF

_findMember:= _findItem(Member, _Item, Result);

IF NOT _findMember		THEN	RETURN;	END_IF
IF _Item = 0 					THEN	RETURN;	END_IF

FoundMember:= _Item^.Member;
END_METHOD

//find a modul by index  
METHOD PROTECTED _findMemberByIndex : BOOL
VAR_INPUT
	Index				: UDINT;	//index of item
	FoundMember	: REFERENCE TO KOSTAL_AF2024_Core_Settings.T_MaxString_UTF8;	//return value
	Result			: KOSTAL_AF2024_Core_functionResponse.I_T_functionResponse_Owner;	//result information
END_VAR

VAR
	_FoundItem	: P_String_UTF8;
END_VAR

IF NOT __ISVALIDREF(FoundMember)	THEN _setResultFail(Result, "FoundMember has no valid reference");	RETURN;	END_IF

FoundMember:= '';

_findMemberByIndex:= _findItemByIndex(Index,_FoundItem, Result);

IF NOT _findMemberByIndex THEN RETURN;	END_IF
IF _FoundItem = 0 THEN RETURN;	END_IF

FoundMember:= _FoundItem^.Member;

_findMemberByIndex:= TRUE;
END_METHOD

METHOD PROTECTED _insertMember : BOOL
VAR_INPUT
	Index		: UDINT;	//Index a which shall inserted the {Item}
	Member	: KOSTAL_AF2024_Core_Settings.T_MaxString_UTF8;
	Result	: KOSTAL_AF2024_Core_functionResponse.I_T_functionResponse_Owner;
END_VAR

VAR
	_Member: KOSTAL_AF2024_Core_System.I_Interface;
END_VAR

_insertMember:= _insertItem(Index, Member, Result);
END_METHOD

(*
	remove Item from begin of list
*)
METHOD PROTECTED _removeFromBegin : BOOL
VAR_INPUT
	Result	: KOSTAL_AF2024_Core_functionResponse.I_T_functionResponse_Owner;
END_VAR

_removeFromBegin:= _removeMemberByIndex(0, Result);
END_METHOD

(*
	remove Item from end of list
*)
METHOD PROTECTED _removeFromEnd : BOOL
VAR_INPUT
	Result	: KOSTAL_AF2024_Core_functionResponse.I_T_functionResponse_Owner;
END_VAR

_removeFromEnd:= _removeMemberByIndex(_Count - 1, Result);
END_METHOD

(*
	remove given {Member} from List
*)
METHOD PROTECTED _removeMember : BOOL
VAR_INPUT
	Member	: KOSTAL_AF2024_Core_Settings.T_MaxString_UTF8;
	Result	: KOSTAL_AF2024_Core_functionResponse.I_T_functionResponse_Owner;
END_VAR

VAR
	_Item		: P_String_UTF8;
	_bFound: BOOL;
END_VAR


_bFound:= _findItem(Member, _Item, Result);

IF NOT _bFound THEN RETURN;	END_IF

_removeMember:= _removeItem(_Item, Result);
END_METHOD

(*
	remove given {Index} from List
*)
METHOD PROTECTED _removeMemberByIndex : BOOL
VAR_INPUT
	Index		: UDINT;
	Result	: KOSTAL_AF2024_Core_functionResponse.I_T_functionResponse_Owner;
END_VAR

VAR
	_bFound	: BOOL;
	_Member	: KOSTAL_AF2024_Core_Settings.T_MaxString_UTF8;

END_VAR

IF NOT _findMemberByIndex(Index, _Member, Result)	THEN RETURN;	END_IF

_removeMemberByIndex:= _removeMember(_Member, Result);
END_METHOD

(*
	Delete the complete content of the list
*)
METHOD PROTECTED _clear
VAR_INPUT
END_VAR

WHILE THIS^._pBegin <> 0 DO
    _removeMember(_pBegin^.Member, 0);  
END_WHILE
END_METHOD

METHOD FB_exit : BOOL
VAR_INPUT
	bInCopyCode : BOOL; // if TRUE, the exit method is called for exiting an instance that is copied afterwards (online change).
END_VAR

_clear();
END_METHOD

METHOD FB_init : BOOL
VAR_INPUT
	bInitRetains : BOOL; // if TRUE, the retain variables are initialized (warm start / cold start)
	bInCopyCode : BOOL;  // if TRUE, the instance afterwards gets moved into the copy code (online change)
END_VAR

_clear();
END_METHOD

END_FUNCTION_BLOCK

// _STRING_UTF8/1_Base/_I_String_UTF8_Base
INTERFACE _I_String_UTF8_Base EXTENDS _I_String_UTF8_Core

END_INTERFACE

// _STRING_UTF8/1_Base/_I_String_UTF8_Base_Owner
INTERFACE _I_String_UTF8_Base_Owner EXTENDS _I_String_UTF8_Core_Owner

END_INTERFACE

// _STRING_UTF8/FB_ListOfString_UTF8
(*
	List of String
	HP -High Performance
	The temporary load on the router's memory is halved.
*)
FUNCTION_BLOCK PUBLIC FB_ListOfString_UTF8 EXTENDS _FB_String_UTF8_Base IMPLEMENTS I_ListOfString_UTF8, I_ListOfString_UTF8_Owner
VAR
	_maxLine	: UDINT:= UDINT#16#FFFF_FFFF;
END_VAR

(*
Description
===========
| Adds a line to end of the list
| Parameters:
| 	line: STRING(255): Text to add to the list
| Returns false in case line is empty or list is full
*)
METHOD addLine : BOOL
VAR_INPUT
	newLine	: KOSTAL_AF2024_Core_Settings.T_MaxString_UTF8;
END_VAR

VAR
	_fRes: KOSTAL_AF2024_Core_functionResponse.T_functionResponse;
END_VAR

addLine:= _addMember(newLine, _fRes) AND _fRes.success;
END_METHOD

(*
Description
===========
| Clears the list's contents
*)
METHOD clear

_clear();
END_METHOD

(*
Description
===========
| Returns the line at the given index
| Parameters:
| 	numberOfLine: index
*)
METHOD line_GET : KOSTAL_AF2024_Core_Settings.T_MaxString_UTF8
VAR_INPUT
	(*1..numberOfLines_GET()*)
	numberOfLine	: UDINT;
END_VAR

VAR
	_fRes: KOSTAL_AF2024_Core_functionResponse.T_functionResponse;
END_VAR

_findMemberByIndex(NumberOfLine - 1, line_GET, _fRes);
END_METHOD

(*
Description
===========
| Returns the line at the given index
| Parameters:
| 	numberOfLine: index
*)
METHOD line_SET : BOOL
VAR_INPUT
	line	: KOSTAL_AF2024_Core_Settings.T_MaxString_UTF8;
	(*1..numberOfLines_GET()*)
	numberOfLine	: UDINT;
END_VAR

VAR
	_item: P_String_UTF8;
	_fRes: KOSTAL_AF2024_Core_functionResponse.T_functionResponse;
END_VAR

IF NOT SUPER^._findItemByIndex(numberOfLine - 1, _item, _fRes)	THEN RETURN;	END_IF

IF NOT _fRes.success	THEN RETURN;	END_IF

IF _item = 0 THEN RETURN;	END_IF

_item^.Member:= line;

line_SET:= TRUE;
END_METHOD

(*
Description
===========
| **Maximum** number of elements in the list. 
| If the list is full, added lines will be ignored
*)
PROPERTY maxLine : UDINT
GET

maxLine:= _maxLine;
END_GET
SET

_maxLine:= maxLine;
END_SET
END_PROPERTY

PROPERTY PUBLIC NumberOfLines : UDINT
GET

NumberOfLines:= SUPER^._Count;
END_GET
END_PROPERTY

(*
Description
===========
| Remove the line with the given index
| Elements after the index move up one position
| Parameters:
| 	index: line to remove
*)
METHOD removeLine
VAR_INPUT
	(*1..numberOfLines_GET()*)
	numberOfLine	: UDINT;
END_VAR

VAR
	_fRes: KOSTAL_AF2024_Core_functionResponse.T_functionResponse;
END_VAR

_removeMemberByIndex(numberOfLine - 1, _fRes);
END_METHOD

END_FUNCTION_BLOCK

// _STRING_UTF8/I_ListOfString_UTF8
INTERFACE I_ListOfString_UTF8 EXTENDS KOSTAL_AF2024_Core_System.I_Interface

(*
Description
===========
| Returns the line at the given index
| Parameters:
| 	numberOfLine: index
*)
METHOD PUBLIC line_GET : KOSTAL_AF2024_Core_Settings.T_MaxString_UTF8
VAR_INPUT
	numberOfLine	:	UDINT;	//1..numberOfLines_GET()
END_VAR
END_METHOD

(*
Description
===========
| **Maximum** number of elements in the list. 
| If the list is full, added lines will be ignored
*)
PROPERTY maxLine : UDINT
GET
END_GET
END_PROPERTY

PROPERTY PUBLIC NumberOfLines : UDINT
GET
END_GET
END_PROPERTY

END_INTERFACE

// _STRING_UTF8/I_ListOfString_UTF8_Owner
INTERFACE I_ListOfString_UTF8_Owner EXTENDS KOSTAL_AF2024_Core_System.I_Interface

(*
Description
===========
| Adds a line to end of the list
| Parameters:
| 	line: STRING(255): Text to add to the list
| Returns false in case line is empty or list is full
*)

METHOD PUBLIC addLine : BOOL
VAR_INPUT
	newLine	: KOSTAL_AF2024_Core_Settings.T_MaxString_UTF8;
END_VAR
END_METHOD

(*
Description
===========
| Clears the list's contents
*)
METHOD PUBLIC clear
VAR_INPUT
END_VAR
END_METHOD

(*
Description
===========
| Returns the line at the given index
| Parameters:
| 	numberOfLine: index
*)
METHOD PUBLIC line_GET :  KOSTAL_AF2024_Core_Settings.T_MaxString_UTF8
VAR_INPUT
	numberOfLine	:	UDINT;	//1..numberOfLines_GET()
END_VAR
END_METHOD

(*
Description
===========
| Returns the line at the given index
| Parameters:
| 	numberOfLine: index
*)
METHOD PUBLIC line_SET : BOOL
VAR_INPUT
	line	:  KOSTAL_AF2024_Core_Settings.T_MaxString_UTF8;
	numberOfLine	:	UDINT;	//1..numberOfLines_GET()
END_VAR
END_METHOD

(*
Description
===========
| **Maximum** number of elements in the list. 
| If the list is full, added lines will be ignored
*)
PROPERTY PUBLIC maxLine : UDINT
GET
END_GET
SET
END_SET
END_PROPERTY

PROPERTY PUBLIC NumberOfLines : UDINT
GET
END_GET
END_PROPERTY

(*
Description
===========
| Remove the line with the given index
| Elements after the index move up one position
| Parameters:
| 	index: line to remove
*)

METHOD PUBLIC removeLine
VAR_INPUT
	numberOfLine	:	UDINT;	//1..numberOfLines_GET()
END_VAR
END_METHOD

END_INTERFACE

// Project Information/F_GetCompany
// This function has been automatically generated from the project information.
{attribute 'signature_flag' := '1073741824'}
{attribute 'TcGenerated'}
{attribute 'no-analysis'}
FUNCTION F_GetCompany : WSTRING
VAR_INPUT
	
END_VAR

F_GetCompany := "KOSTAL GmbH & Co.KG";

END_FUNCTION

// Project Information/F_GetTitle
// This function has been automatically generated from the project information.
{attribute 'signature_flag' := '1073741824'}
{attribute 'TcGenerated'}
{attribute 'no-analysis'}
FUNCTION F_GetTitle : WSTRING
VAR_INPUT
	
END_VAR

F_GetTitle := "KOSTAL.AF2024.Core.ListOf";

END_FUNCTION

// Project Information/F_GetVersion
// This function has been automatically generated from the project information.
{attribute 'signature_flag' := '1073741824'}
{attribute 'TcGenerated'}
{attribute 'no-analysis'}
FUNCTION F_GetVersion : ST_LibVersion
VAR_INPUT
	
END_VAR

F_GetVersion.iMajor := 1;
F_GetVersion.iMinor := 0;
F_GetVersion.iBuild := 0;
F_GetVersion.iRevision := 0;
F_GetVersion.sVersion := '1.0.0.0';
F_GetVersion.nFlags := 0;

END_FUNCTION
